INTERFACE I_Valve

METHOD Close : BOOL
END_METHOD

METHOD Open : BOOL
VAR_INPUT
	bForce	: BOOL;
END_VAR
END_METHOD

PROPERTY State : E_ValveState
GET // PUBLIC
END_GET
END_PROPERTY

END_INTERFACE

(* stored: Version 1.1.0.1
   Itf I_Valve: Id {b219a1d8-09d2-4b1b-8ade-b912b76d7381}
   Method Close: Id {834bc315-e0a3-4811-b0c5-9d5d3e765d9a}
   Method Open: Id {a373a831-d91e-42b8-af1f-8cf9ff5e8817}
   Property State: Id {5c836057-bd2e-40c5-9d53-654234c8df2d}
   Get Get: Id {26ed08ba-6895-4b64-8545-cecf46e66dc7} *)
